// TIA Portal V21 export
ORGANIZATION_BLOCK "LongNames"   // OB1, LAD
BEGIN

REGION Network 1: Long tag names
   // A comment that runs on.
   // And a second line.
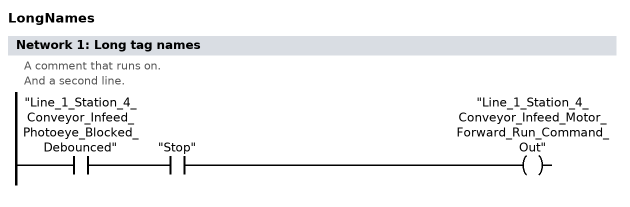
   RUNG wire#powerrail
      Contact( "Line_1_Station_4_Conveyor_Infeed_Photoeye_Blocked_Debounced" )
      Contact( "Stop" )
      Coil( "Line_1_Station_4_Conveyor_Infeed_Motor_Forward_Run_Command_Out" )
   END_RUNG
   // the same network as SCL:
   "Line_1_Station_4_Conveyor_Infeed_Motor_Forward_Run_Command_Out" := "Line_1_Station_4_Conveyor_Infeed_Photoeye_Blocked_Debounced" AND "Stop";
END_REGION
END_ORGANIZATION_BLOCK
